Staubli VAL3: resetBusSelect.pgx

program resetBusSelect(num x_nIndex)
  local num i
begin
  for i =0 to 5
    if i!=x_nIndex
      bBusSelect[i]=false
    endIf
  endFor
end
